(* IEC 61131-3 sources: codesys-framework/txt/application/ToDo/Hardware/IO/Cylinder/DUT, 2 files *)

(* ---- E_CylinderStates.dut.st ---- *)
{attribute 'qualified_only'}
{attribute 'strict'}
TYPE E_CylinderStates :
(
	Invalid := 0,
	Pos0,
	Pos1,
	GoToPos0,
	GoToPos1
);
END_TYPE

(* ---- SC_SystemParametersCylinder.dut.st ---- *)
TYPE SC_SystemParametersCylinder:
STRUCT
	xSensorPresentPos0		: BOOL;
	xSensorPresentPos1		: BOOL;

	xSensorCriticalPos0		: BOOL := TRUE;
	xSensorCriticalPos1		: BOOL := TRUE;

	tCylinderToPos0			: TIME;
	tCylinderToPos1			: TIME;

	rErrorTimeoutFactor		: REAL := 1;
END_STRUCT
END_TYPE
